Staubli VAL3: main.pgx

public program main()
  local num l_j
  local num l_i
begin
  for l_i = 0 to size(aActItem)-1
    aActItem[l_i].sComment="Action"+toString("",l_i)
    for l_j = 0 to size(aActItem[l_i].aActItem)-1
      aActItem[l_i].aActItem[l_j].nIOindex=-1
    endFor

  endFor
  libSave()
end
